(* IEC 61131-3 sources: llm-plc-st-eval/data/processed_definitivo/claude-sonnet-4-6/A3/zero_shot, 3 files *)

(* ---- ejec_1.st ---- *)
FUNCTION_BLOCK FB_Com
VAR_INPUT
    txReq  : BOOL; (* Solicitud de transmisión *)
    rxOk   : BOOL; (* Confirmación de recepción del dispositivo externo *)
    rxData : INT;  (* Dato recibido (eco) *)
END_VAR

VAR_OUTPUT
    txData   : INT;  (* Dato transmitido *)
    ocupado  : BOOL; (* Intercambio en curso *)
    ok       : BOOL; (* Último intercambio exitoso *)
    error    : BOOL; (* Fallaron los 3 intentos *)
    nIntentos: INT;  (* Número de intento en curso / último *)
END_VAR

VAR
    txReq_prev : BOOL;        (* Valor anterior de txReq para detectar flanco *)
    timer      : TON;         (* Temporizador de plazo por intento *)
    timerRun   : BOOL;        (* Habilita el temporizador *)
    TEST_VALUE : INT := 100;  (* Valor de prueba fijo *)
    MAX_INT    : INT := 3;    (* Máximo número de intentos *)
END_VAR

(* ── Temporizador ── *)
timer(IN := timerRun, PT := T#500MS);

(* ── Detección de flanco ascendente en txReq ── *)
IF txReq AND NOT txReq_prev THEN
    IF NOT ocupado THEN
        (* Iniciar nuevo intercambio *)
        ok        := FALSE;
        error     := FALSE;
        ocupado   := TRUE;
        nIntentos := 1;
        txData    := TEST_VALUE;
        timerRun  := TRUE;   (* Arrancar temporizador del intento 1 *)
    END_IF;
    (* Si ocupado = TRUE, el flanco se ignora *)
END_IF;

(* ── Lógica principal durante un intercambio ── *)
IF ocupado THEN

    IF rxOk THEN
        (* Ha llegado respuesta del dispositivo *)
        IF rxData = txData THEN
            (* ── Intento correcto ── *)
            timerRun := FALSE;
            ocupado  := FALSE;
            ok       := TRUE;
        ELSE
            (* ── Respuesta incorrecta: tratar como fallo de intento ── *)
            timerRun := FALSE;          (* Detener y resetear temporizador *)
            IF nIntentos < MAX_INT THEN
                nIntentos := nIntentos + 1;
                timerRun  := TRUE;      (* Nuevo plazo para el siguiente intento *)
            ELSE
                (* Agotados los 3 intentos *)
                ocupado := FALSE;
                error   := TRUE;
            END_IF;
        END_IF;

    ELSIF timer.Q THEN
        (* ── Plazo vencido sin confirmación ── *)
        timerRun := FALSE;              (* Resetear temporizador *)
        IF nIntentos < MAX_INT THEN
            nIntentos := nIntentos + 1;
            timerRun  := TRUE;          (* Nuevo plazo para el siguiente intento *)
        ELSE
            (* Agotados los 3 intentos *)
            ocupado := FALSE;
            error   := TRUE;
        END_IF;
    END_IF;

END_IF;

(* ── Guardar estado anterior de txReq ── *)
txReq_prev := txReq;

(* ---- ejec_2.st ---- *)
FUNCTION_BLOCK FB_Com

VAR_INPUT
    txReq  : BOOL; (* Solicitud de transmisión *)
    rxOk   : BOOL; (* Confirmación de recepción del dispositivo externo *)
    rxData : INT;  (* Dato recibido (eco) *)
END_VAR

VAR_OUTPUT
    txData   : INT;  (* Dato transmitido *)
    ocupado  : BOOL; (* Intercambio en curso *)
    ok       : BOOL; (* Último intercambio correcto *)
    error    : BOOL; (* Fallaron los 3 intentos *)
    nIntentos: INT;  (* Número de intento en curso / último *)
END_VAR

VAR
    txReq_prev : BOOL;        (* Valor anterior de txReq para detectar flanco *)
    timer      : TON;         (* Temporizador de 500 ms por intento *)
    timerStart : BOOL;        (* Señal de arranque del temporizador *)
    TEST_VALUE : INT := 100;  (* Valor de prueba fijo *)
    MAX_INTENTOS : INT := 3;  (* Máximo de intentos permitidos *)
END_VAR

(* ─────────────────────────────────────────────────────────────
   Detección de flanco ascendente en txReq
   ───────────────────────────────────────────────────────────── *)
IF txReq AND NOT txReq_prev THEN
    (* Flanco detectado: iniciar intercambio solo si no hay uno en curso *)
    IF NOT ocupado THEN
        ocupado   := TRUE;
        ok        := FALSE;
        error     := FALSE;
        nIntentos := 1;
        txData    := TEST_VALUE;
        timerStart := FALSE; (* Forzar reinicio del TON en el siguiente ciclo *)
    END_IF;
END_IF;
txReq_prev := txReq;

(* ─────────────────────────────────────────────────────────────
   Lógica principal: solo activa cuando hay intercambio en curso
   ───────────────────────────────────────────────────────────── *)
IF ocupado THEN

    (* Arrancar / mantener el temporizador del intento actual *)
    timerStart := TRUE;
    timer(IN := timerStart, PT := T#500MS);

    (* Comprobar respuesta correcta: rxOk activo y eco coincide *)
    IF rxOk AND (rxData = txData) THEN
        (* Intento exitoso *)
        ok        := TRUE;
        ocupado   := FALSE;
        timerStart := FALSE;
        timer(IN := FALSE, PT := T#500MS); (* Detener temporizador *)

    (* Comprobar fallo: tiempo agotado O rxOk con dato incorrecto *)
    ELSIF timer.Q OR (rxOk AND (rxData <> txData)) THEN
        (* Intento fallido *)
        IF nIntentos < MAX_INTENTOS THEN
            (* Iniciar siguiente intento *)
            nIntentos  := nIntentos + 1;
            timerStart := FALSE;             (* Bajar IN para reiniciar TON *)
            timer(IN := FALSE, PT := T#500MS);
            (* timerStart se volverá TRUE en el próximo ciclo *)
        ELSE
            (* Se agotaron los 3 intentos *)
            error      := TRUE;
            ocupado    := FALSE;
            timerStart := FALSE;
            timer(IN := FALSE, PT := T#500MS); (* Detener temporizador *)
        END_IF;
    END_IF;

END_IF;

(* Llamada final al temporizador para actualizar su salida Q *)
timer(IN := timerStart, PT := T#500MS);

(* ---- ejec_3.st ---- *)
FUNCTION_BLOCK FB_Com
VAR_INPUT
    txReq  : BOOL; (* Solicitud de transmisión *)
    rxOk   : BOOL; (* Confirmación de recepción del dispositivo externo *)
    rxData : INT;  (* Dato recibido (eco) *)
END_VAR

VAR_OUTPUT
    txData   : INT;  (* Dato transmitido *)
    ocupado  : BOOL; (* Intercambio en curso *)
    ok       : BOOL; (* Último intercambio exitoso *)
    error    : BOOL; (* Fallaron los 3 intentos *)
    nIntentos: INT;  (* Número de intento en curso / último intento realizado *)
END_VAR

VAR
    txReq_prev : BOOL;       (* Valor anterior de txReq para detectar flanco ascendente *)
    timer      : TON;        (* Temporizador de plazo por intento *)
    activo     : BOOL;       (* Intercambio en curso internamente *)
    valorTx    : INT := 100; (* Valor de prueba fijo *)
END_VAR

(* ── Detección de flanco ascendente de txReq ── *)
IF txReq AND NOT txReq_prev THEN
    IF NOT activo THEN
        (* Iniciar nuevo intercambio *)
        activo    := TRUE;
        ocupado   := TRUE;
        ok        := FALSE;
        error     := FALSE;
        nIntentos := 1;
        txData    := valorTx;
        (* Arrancar temporizador del primer intento *)
        timer(IN := FALSE, PT := T#500MS);
        timer(IN := TRUE,  PT := T#500MS);
    END_IF;
    (* Si activo = TRUE, el flanco se ignora *)
END_IF;

(* ── Lógica principal del intercambio ── *)
IF activo THEN
    (* Actualizar temporizador *)
    timer(IN := TRUE, PT := T#500MS);

    (* Comprobar respuesta correcta: rxOk activo y eco coincide *)
    IF rxOk AND (rxData = txData) THEN
        (* Intento exitoso *)
        ok      := TRUE;
        error   := FALSE;
        ocupado := FALSE;
        activo  := FALSE;
        timer(IN := FALSE, PT := T#500MS); (* Detener temporizador *)

    (* Comprobar fallo: plazo vencido O rxOk con dato incorrecto *)
    ELSIF timer.Q OR (rxOk AND (rxData <> txData)) THEN
        (* Intento fallido *)
        timer(IN := FALSE, PT := T#500MS); (* Resetear temporizador *)

        IF nIntentos < 3 THEN
            (* Iniciar siguiente intento *)
            nIntentos := nIntentos + 1;
            txData    := valorTx;
            timer(IN := TRUE, PT := T#500MS); (* Arrancar nuevo plazo *)
        ELSE
            (* Agotados los 3 intentos *)
            error   := TRUE;
            ok      := FALSE;
            ocupado := FALSE;
            activo  := FALSE;
        END_IF;
    END_IF;
END_IF;

(* ── Guardar estado anterior de txReq ── *)
txReq_prev := txReq;
